// TIA Portal V21 export
// export: Created 2026-11-11T00:49:03.0617986Z, ExportSetting WithDefaults, DisplayName Totally Integrated Automation Portal, DisplayVersion V21 Update 3, DisplayName STEP 7 Professional, DisplayVersion V21 Update 3, DisplayName STEP 7 Safety, DisplayVersion V21, DisplayName Tech WebApplication, DisplayVersion V21, DisplayName WinCC Basic/Comfort/Advanced, DisplayVersion V21 Update 3, DisplayName WinCC Unified, DisplayVersion V21 Update 3
FUNCTION_BLOCK "FX_Lad_ex093"   // FB231, LAD
{ S7_Optimized_Access := 'TRUE' }
VERSION : 0.1
// stored: AutoNumber true, IsIECCheckEnabled false, IsRetainMemResEnabled false, MemoryReserve 100, SetENOAutomatically false, UDAEnableTagReadback false
   VAR_INPUT
      "a" : Bool;
      "b" : Bool;
      c : Bool;
      ia : Int;
      ib : Int;
      ic : Int;
      da : DInt;
      db : DInt;
      ra : Real;
      rb : Real;
      wa : Word;
      wb : Word;
      dwa : DWord;
      ba : Byte;
      ta : Time;
      tb : Time;
      s1 : String;
      s2 : String;
   END_VAR
   VAR_OUTPUT
      q : Bool;
      q2 : Bool;
      io : Int;
      io2 : Int;
      dout : DInt;
      rout : Real;
      wout : Word;
      dwout : DWord;
      bout : Byte;
      tout : Time;
      sout : String;
   END_VAR
   VAR_IN_OUT
      p_pe_i_dev_new : Bool;
      p_cmd : Int;
      p_start_pause : Bool;
      p_activate : Bool;
      p_valid : Bool;
      p_error : Bool;
      p_status : Word;
      arr : Array[0..9] of Int;
      barr : Array[0..7] of Bool;
      iinout : Int;
   END_VAR
   VAR
      ton1 { S7_SetPoint := 'True'} : TON_TIME;
      tof1 { S7_SetPoint := 'True'} : TOF_TIME;
      tp1 { S7_SetPoint := 'True'} : TP_TIME;
      tonr1 { S7_SetPoint := 'True'} : TONR_TIME;
      ctu1 { S7_SetPoint := 'True'} : CTU_INT;
      ctd1 { S7_SetPoint := 'True'} : CTD_INT;
      ctud1 { S7_SetPoint := 'True'} : CTUD_INT;
      rtrig1 { S7_SetPoint := 'True'} : R_TRIG;
      ftrig1 { S7_SetPoint := 'True'} : F_TRIG;
      edge1 : Bool;
      edge2 : Bool;
      stat1 : Bool;
      stat2 : Bool;
      stati : Int;
   END_VAR
   VAR_TEMP
      t1 : Bool;
      t2 : Bool;
      ti : Int;
      td : DInt;
      tr : Real;
      tw : Word;
      tt : Time;
      var1 : Variant;
   END_VAR
BEGIN

REGION Network 1: ---| |--- - Normally open contact
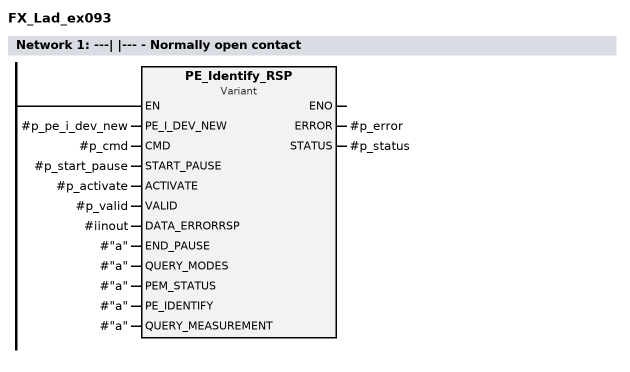
   RUNG wire#powerrail
      { S7_Templates := "data_errorrsp_type := Variant" } PE_Identify_RSP(PE_I_DEV_NEW := #p_pe_i_dev_new, CMD := #p_cmd, Start_Pause := #p_start_pause, Activate := #p_activate, VALID := #p_valid, DATA_ERRORRSP := #iinout, ERROR => #p_error, STATUS => #p_status, End_Pause := #"a", Query_Modes := #"a", PEM_Status := #"a", PE_Identify := #"a", Query_Measurement := #"a")
   END_RUNG
   // the same network as SCL:
   PE_Identify_RSP(PE_I_DEV_NEW := #p_pe_i_dev_new,
                   CMD := #p_cmd,
                   Start_Pause := #p_start_pause,
                   Activate := #p_activate,
                   VALID := #p_valid,
                   DATA_ERRORRSP := #iinout,
                   End_Pause := #"a",
                   Query_Modes := #"a",
                   PEM_Status := #"a",
                   PE_Identify := #"a",
                   Query_Measurement := #"a",
                   ERROR => #p_error,
                   STATUS => #p_status);
END_REGION
END_FUNCTION_BLOCK
